(* IEC 61131-3 sources: llm-plc-st-eval/data/definitivo/gpt-4o-2024-08-06/I5/few_shot, 3 files *)

(* ---- ejec_1.st ---- *)
```pascal
FUNCTION_BLOCK FB_Clasificadora
VAR_INPUT
    sensorPresencia : BOOL; (* Sensor de presencia de piezas *)
    sensorAltura : BOOL;    (* Sensor de altura de piezas *)
END_VAR
VAR_OUTPUT
    banda : BOOL;           (* Banda transportadora activa *)
    piston : BOOL;          (* Pistón para desviar piezas altas *)
    nAltas : INT;           (* Contador de piezas altas *)
    nBajas : INT;           (* Contador de piezas bajas *)
END_VAR
VAR
    tRetraso : TON;         (* Temporizador de retraso de 2 segundos *)
    tPulso : TON;           (* Temporizador de pulso de 1 segundo *)
    piezaAltaDetectada : BOOL; (* Indica si una pieza alta fue detectada *)
END_VAR

(* La banda transportadora siempre está activa *)
banda := TRUE;

(* Detectar y contar piezas *)
IF sensorPresencia THEN
    IF sensorAltura THEN
        nAltas := nAltas + 1;
        piezaAltaDetectada := TRUE;
        tRetraso(IN := TRUE, PT := T#2S);
    ELSE
        nBajas := nBajas + 1;
    END_IF;
END_IF;

(* Control del pistón para desviar piezas altas *)
IF piezaAltaDetectada AND tRetraso.Q THEN
    tPulso(IN := TRUE, PT := T#1S);
    piezaAltaDetectada := FALSE; (* Resetear la detección de pieza alta *)
END_IF;

piston := tPulso.Q;
END_FUNCTION_BLOCK
```

(* ---- ejec_2.st ---- *)
```pascal
FUNCTION_BLOCK FB_Clasificadora
VAR_INPUT
    sensorPresencia : BOOL; (* Sensor de presencia de piezas *)
    sensorAltura : BOOL;    (* Sensor de altura de piezas *)
END_VAR
VAR_OUTPUT
    banda : BOOL;           (* Banda transportadora activa *)
    piston : BOOL;          (* Pistón para desviar piezas altas *)
    nAltas : INT;           (* Contador de piezas altas *)
    nBajas : INT;           (* Contador de piezas bajas *)
END_VAR
VAR
    tRetraso : TON;         (* Temporizador para retraso de 2 segundos *)
    tPulso : TP;            (* Temporizador para pulso de 1 segundo *)
    piezaAltaDetectada : BOOL; (* Indica si una pieza alta fue detectada *)
END_VAR

(* La banda transportadora siempre está activa *)
banda := TRUE;

(* Detectar y contar piezas altas y bajas *)
IF sensorPresencia THEN
    IF sensorAltura THEN
        (* Si la pieza es alta, incrementar el contador de piezas altas *)
        nAltas := nAltas + 1;
        piezaAltaDetectada := TRUE;
        tRetraso(IN := TRUE, PT := T#2S);
    ELSE
        (* Si la pieza es baja, incrementar el contador de piezas bajas *)
        nBajas := nBajas + 1;
    END_IF;
END_IF;

(* Activar el pistón después de 2 segundos si una pieza alta fue detectada *)
IF tRetraso.Q THEN
    tPulso(IN := piezaAltaDetectada, PT := T#1S);
    piezaAltaDetectada := FALSE; (* Resetear la detección de pieza alta *)
END_IF;

(* Salida del pistón activada por el pulso de 1 segundo *)
piston := tPulso.Q;
END_FUNCTION_BLOCK
```

(* ---- ejec_3.st ---- *)
```pascal
FUNCTION_BLOCK FB_Clasificadora
VAR_INPUT
    sensorPresencia : BOOL; (* Sensor de presencia de piezas *)
    sensorAltura : BOOL;    (* Sensor de altura de piezas *)
END_VAR
VAR_OUTPUT
    banda : BOOL;   (* Banda transportadora activa *)
    piston : BOOL;  (* Pistón para desviar piezas altas *)
    nAltas : INT;   (* Contador de piezas altas *)
    nBajas : INT;   (* Contador de piezas bajas *)
END_VAR
VAR
    tRetraso : TON; (* Temporizador para retraso de 2 segundos *)
    tPiston : TON;  (* Temporizador para activación de pistón por 1 segundo *)
    piezaAltaDetectada : BOOL; (* Indica si una pieza alta fue detectada *)
END_VAR

(* La banda siempre está activa *)
banda := TRUE;

(* Detectar y contar piezas *)
IF sensorPresencia THEN
    IF sensorAltura THEN
        nAltas := nAltas + 1;
        piezaAltaDetectada := TRUE;
        tRetraso(IN := TRUE, PT := T#2S);
    ELSE
        nBajas := nBajas + 1;
    END_IF;
END_IF;

(* Control del pistón *)
IF tRetraso.Q THEN
    tPiston(IN := piezaAltaDetectada, PT := T#1S);
    piezaAltaDetectada := FALSE; (* Resetear la detección de pieza alta después del retraso *)
END_IF;

piston := tPiston.Q;
END_FUNCTION_BLOCK
```
